// TwinCAT 3 PLC project TcoCognexVisionTests
// Title: TcoCognexVisionTests
// Company: Vortex.Library
// ProjectVersion: 0.6.0.913
// ProgramVersion: 3.1.4024.12
// libraries:
//   Tc2_Standard, * (Beckhoff Automation GmbH)
//   Tc2_System, * (Beckhoff Automation GmbH)
//   Tc3_Module, * (Beckhoff Automation GmbH)
//   TcoAbstractions, 0.6.0.913 (Vortex.Library)
//   TcoCognexVision, 0.6.0.913 (Vortex.Library)
//   TcoCore, 0.6.0.913 (Vortex.Library)
//   TcoInspectors, 0.6.0.913 (Vortex.Library)
//   TcoIo, 0.6.0.913 (Vortex.Library)
//   TcoUtilities, 0.6.0.913 (Vortex.Library)
// project tree:
//   DUTs/ DesignerResults.TcDUT, DesignerUserData.TcDUT
//   GVLs/ GVL.TcGVL
//   / PlcTask.TcTTO
//   POUs/ ITcoResultsData.TcIO, MAIN.TcPOU, myVeryFirstTcoContext.TcPOU, ProjectSpecificData.TcPOU
// (motion and I/O tree: see PLC project tcocognexvision)
// real-time tasks:
//   TASK PlcTask: cycle T#10ms, priority 20, ADS port 350
//   TASK PNIO: cycle T#16ms, priority 21, ADS port 351
//   TASK PlcTask1: cycle T#10ms, priority 22, ADS port 352
// variable links:
//   TcoCognexVisionTests/TcoCognexVisionTests Instance <-> Device 1 (Profinet Controller)/myveryfirstdataman
//     PlcTask Inputs/GVL.myVeryFirstDatamanGVL.AcquisitionStatus.Acquiring <-> API/Acquisition_Status/Acquisition_Status/Inputs/Acquisition_Status_Register/Acquiring
//     PlcTask Inputs/GVL.myVeryFirstDatamanGVL.AcquisitionStatus.MissedAcquisition <-> API/Acquisition_Status/Acquisition_Status/Inputs/Acquisition_Status_Register/Missed_Acquisition
//     PlcTask Inputs/GVL.myVeryFirstDatamanGVL.AcquisitionStatus.TriggerAcknowledge <-> API/Acquisition_Status/Acquisition_Status/Inputs/Acquisition_Status_Register/Trigger_Acknowledge
//     PlcTask Inputs/GVL.myVeryFirstDatamanGVL.AcquisitionStatus.TriggerID <-> API/Acquisition_Status/Acquisition_Status/Inputs/Trigger_ID
//     PlcTask Inputs/GVL.myVeryFirstDatamanGVL.AcquisitionStatus.TriggerReady <-> API/Acquisition_Status/Acquisition_Status/Inputs/Acquisition_Status_Register/Trigger_Ready
//     PlcTask Inputs/GVL.myVeryFirstDatamanGVL.PnIoBoxDiag <-> Inputs/PnIoBoxDiag
//     PlcTask Inputs/GVL.myVeryFirstDatamanGVL.PnIoBoxState <-> Inputs/PnIoBoxState
//     PlcTask Inputs/GVL.myVeryFirstDatamanGVL.ResultData.ResultCode <-> API/Result_Data_64_bytes/Result_Data_64_bytes/Inputs/Result_Code
//     PlcTask Inputs/GVL.myVeryFirstDatamanGVL.ResultData.ResultData <-> API/Result_Data_64_bytes/Result_Data_64_bytes/Inputs/Result_Data
//     PlcTask Inputs/GVL.myVeryFirstDatamanGVL.ResultData.ResultExtended <-> API/Result_Data_64_bytes/Result_Data_64_bytes/Inputs/Result_Extended
//     PlcTask Inputs/GVL.myVeryFirstDatamanGVL.ResultData.ResultID <-> API/Result_Data_64_bytes/Result_Data_64_bytes/Inputs/Result_ID
//     PlcTask Inputs/GVL.myVeryFirstDatamanGVL.ResultData.ResultLength <-> API/Result_Data_64_bytes/Result_Data_64_bytes/Inputs/Result_Length
//     PlcTask Inputs/GVL.myVeryFirstDatamanGVL.ResultsStatus.DecodeComplete <-> API/Results_Status/Results_Status/Inputs/Results_Status_Register/Decode_Complete
//     PlcTask Inputs/GVL.myVeryFirstDatamanGVL.ResultsStatus.Decoding <-> API/Results_Status/Results_Status/Inputs/Results_Status_Register/Decoding
//     PlcTask Inputs/GVL.myVeryFirstDatamanGVL.ResultsStatus.ErrorDetected <-> API/Results_Status/Results_Status/Inputs/Results_Status_Register/Set_when_reader_fault_occurs
//     PlcTask Inputs/GVL.myVeryFirstDatamanGVL.ResultsStatus.ResultsAvailable <-> API/Results_Status/Results_Status/Inputs/Results_Status_Register/Results_Available
//     PlcTask Inputs/GVL.myVeryFirstDatamanGVL.ResultsStatus.ResultsBufferOverrun <-> API/Results_Status/Results_Status/Inputs/Results_Status_Register/Results_Buffer_Overrun
//     PlcTask Inputs/GVL.myVeryFirstDatamanGVL.SoftEventControl.ExecuteDMCCAcknowledge <-> API/Soft_Event_Control/Soft_Event_Control/Inputs/Soft_Event_Acknowledge_Register/Execute_DMCC_Acknowledge
//     PlcTask Inputs/GVL.myVeryFirstDatamanGVL.SoftEventControl.SetMatchStringAcknowledge <-> API/Soft_Event_Control/Soft_Event_Control/Inputs/Soft_Event_Acknowledge_Register/Set_Match_String_Acknowledge
//     PlcTask Inputs/GVL.myVeryFirstDatamanGVL.SoftEventControl.TrainBrightnessAcknowledge <-> API/Soft_Event_Control/Soft_Event_Control/Inputs/Soft_Event_Acknowledge_Register/Train_Brightness_Acknowledge
//     PlcTask Inputs/GVL.myVeryFirstDatamanGVL.SoftEventControl.TrainCodeAcknowledge <-> API/Soft_Event_Control/Soft_Event_Control/Inputs/Soft_Event_Acknowledge_Register/Train_Code_Acknowledge
//     PlcTask Inputs/GVL.myVeryFirstDatamanGVL.SoftEventControl.TrainFocusAcknowledge <-> API/Soft_Event_Control/Soft_Event_Control/Inputs/Soft_Event_Acknowledge_Register/Train_Focus_Acknowledge
//     PlcTask Inputs/GVL.myVeryFirstDatamanGVL.SoftEventControl.TrainMatchStringAcknowledge <-> API/Soft_Event_Control/Soft_Event_Control/Inputs/Soft_Event_Acknowledge_Register/Train_Match_String_Acknowledge
//     PlcTask Inputs/GVL.myVeryFirstDatamanGVL.SoftEventControl.UntrainAcknowledge <-> API/Soft_Event_Control/Soft_Event_Control/Inputs/Soft_Event_Acknowledge_Register/Untrain_Acknowledge
//     PlcTask Outputs/GVL.myVeryFirstDatamanGVL.AcquisitionControl.Trigger <-> API/Acquisition_Control/Acquisition_Control/Outputs/Acquisition_Control_Register/Trigger
//     PlcTask Outputs/GVL.myVeryFirstDatamanGVL.AcquisitionControl.TriggerEnable <-> API/Acquisition_Control/Acquisition_Control/Outputs/Acquisition_Control_Register/Trigger_Enable
//     PlcTask Outputs/GVL.myVeryFirstDatamanGVL.PnIoBoxCtrl <-> Outputs/PnIoBoxCtrl
//     PlcTask Outputs/GVL.myVeryFirstDatamanGVL.ResultsControl.EnableResultBuffering <-> API/Results_Control/Results_Control/Outputs/Results_Control_Register/Enable_Result_Buffering
//     PlcTask Outputs/GVL.myVeryFirstDatamanGVL.ResultsControl.ResultsAcknowledge <-> API/Results_Control/Results_Control/Outputs/Results_Control_Register/Results_Acknowledge
//     PlcTask Outputs/GVL.myVeryFirstDatamanGVL.SoftEventControl.ExecuteDMCC <-> API/Soft_Event_Control/Soft_Event_Control/Outputs/Soft_Event_Control_Register/Execute_DMCC
//     PlcTask Outputs/GVL.myVeryFirstDatamanGVL.SoftEventControl.SetMatchString <-> API/Soft_Event_Control/Soft_Event_Control/Outputs/Soft_Event_Control_Register/Set_Match_String
//     PlcTask Outputs/GVL.myVeryFirstDatamanGVL.SoftEventControl.TrainBrightness <-> API/Soft_Event_Control/Soft_Event_Control/Outputs/Soft_Event_Control_Register/Train_Brightness
//     PlcTask Outputs/GVL.myVeryFirstDatamanGVL.SoftEventControl.TrainCode <-> API/Soft_Event_Control/Soft_Event_Control/Outputs/Soft_Event_Control_Register/Train_Code
//     PlcTask Outputs/GVL.myVeryFirstDatamanGVL.SoftEventControl.TrainFocus <-> API/Soft_Event_Control/Soft_Event_Control/Outputs/Soft_Event_Control_Register/Train_Focus
//     PlcTask Outputs/GVL.myVeryFirstDatamanGVL.SoftEventControl.TrainMatchString <-> API/Soft_Event_Control/Soft_Event_Control/Outputs/Soft_Event_Control_Register/Train_Match_String
//     PlcTask Outputs/GVL.myVeryFirstDatamanGVL.SoftEventControl.Untrain <-> API/Soft_Event_Control/Soft_Event_Control/Outputs/Soft_Event_Control_Register/Untrain
//     PlcTask Outputs/GVL.myVeryFirstDatamanGVL.UserData.UserData <-> API/User_Data_64_bytes/User_Data_64_bytes/Outputs/User_Data
//     PlcTask Outputs/GVL.myVeryFirstDatamanGVL.UserData.UserDataLength <-> API/User_Data_64_bytes/User_Data_64_bytes/Outputs/User_Data_Length
//     PlcTask Outputs/GVL.myVeryFirstDatamanGVL.UserData.UserDataOption <-> API/User_Data_64_bytes/User_Data_64_bytes/Outputs/User_Data_Option
//   TcoCognexVisionTests/TcoCognexVisionTests Instance <-> Device 1 (Profinet Controller)/myveryfirstinsight
//     PlcTask Inputs/GVL.myVeryFirstInsightGVL.AcquisitionStatus.AcquisitionID <-> API/Acquisition_Status/Acquisition_Status/Inputs/Acquisition_ID
//     PlcTask Inputs/GVL.myVeryFirstInsightGVL.AcquisitionStatus.AcquisitionTriggerAcknowledge <-> API/Acquisition_Status/Acquisition_Status/Inputs/Acquisition_Status_Register/Acquisition_Trigger_Acknowledge
//     PlcTask Inputs/GVL.myVeryFirstInsightGVL.AcquisitionStatus.AcquisitionTriggerReady <-> API/Acquisition_Status/Acquisition_Status/Inputs/Acquisition_Status_Register/Acquisition_Trigger_Ready
//     PlcTask Inputs/GVL.myVeryFirstInsightGVL.AcquisitionStatus.ExposureComplete <-> API/Acquisition_Status/Acquisition_Status/Inputs/Acquisition_Status_Register/Exposure_Complete
//     PlcTask Inputs/GVL.myVeryFirstInsightGVL.AcquisitionStatus.MissedAcquisition <-> API/Acquisition_Status/Acquisition_Status/Inputs/Acquisition_Status_Register/Missed_Acquisition
//     PlcTask Inputs/GVL.myVeryFirstInsightGVL.AcquisitionStatus.OfflineReason0 <-> API/Acquisition_Status/Acquisition_Status/Inputs/Acquisition_Status_Register/Offline_Reason_0
//     PlcTask Inputs/GVL.myVeryFirstInsightGVL.AcquisitionStatus.OfflineReason1 <-> API/Acquisition_Status/Acquisition_Status/Inputs/Acquisition_Status_Register/Offline_Reason_1
//     PlcTask Inputs/GVL.myVeryFirstInsightGVL.AcquisitionStatus.OfflineReason2 <-> API/Acquisition_Status/Acquisition_Status/Inputs/Acquisition_Status_Register/Offline_Reason_2
//     PlcTask Inputs/GVL.myVeryFirstInsightGVL.AcquisitionStatus.Online <-> API/Acquisition_Status/Acquisition_Status/Inputs/Acquisition_Status_Register/Online
//     PlcTask Inputs/GVL.myVeryFirstInsightGVL.CommandControl.CurrentJobID <-> API/Command_Control/Command_Control/Inputs/Current_Job_ID
//     PlcTask Inputs/GVL.myVeryFirstInsightGVL.InspectionStatus.CommandComplete <-> API/Inspection_Status/Inspection_Status/Inputs/Inspection_Status_Register/Command_Complete
//     PlcTask Inputs/GVL.myVeryFirstInsightGVL.InspectionStatus.CommandExecuting <-> API/Inspection_Status/Inspection_Status/Inputs/Inspection_Status_Register/Command_Executing
//     PlcTask Inputs/GVL.myVeryFirstInsightGVL.InspectionStatus.CommandFailed <-> API/Inspection_Status/Inspection_Status/Inputs/Inspection_Status_Register/Command_Failed
//     PlcTask Inputs/GVL.myVeryFirstInsightGVL.InspectionStatus.Error <-> API/Inspection_Status/Inspection_Status/Inputs/Inspection_Status_Register/Error
//     PlcTask Inputs/GVL.myVeryFirstInsightGVL.InspectionStatus.ErrorCode <-> API/Inspection_Status/Inspection_Status/Inputs/Error_Code
//     PlcTask Inputs/GVL.myVeryFirstInsightGVL.InspectionStatus.ExtendedUserDataSetAcknowledge <-> API/Inspection_Status/Inspection_Status/Inputs/Inspection_Status_Register/Extended_User_Data_Set_Acknowledge
//     PlcTask Inputs/GVL.myVeryFirstInsightGVL.InspectionStatus.InspectionCompleted <-> API/Inspection_Status/Inspection_Status/Inputs/Inspection_Status_Register/Inspection_Completed
//     PlcTask Inputs/GVL.myVeryFirstInsightGVL.InspectionStatus.OverallJobPassFail <-> API/Inspection_Status/Inspection_Status/Inputs/Inspection_Status_Register/Set_when_last_inspection_passed,_based_on_the_Overall_Job_Pass_Fail_cell
//     PlcTask Inputs/GVL.myVeryFirstInsightGVL.InspectionStatus.ResultsBufferOverrun <-> API/Inspection_Status/Inspection_Status/Inputs/Inspection_Status_Register/Results_Buffer_Overrun
//     PlcTask Inputs/GVL.myVeryFirstInsightGVL.InspectionStatus.ResultsValid <-> API/Inspection_Status/Inspection_Status/Inputs/Inspection_Status_Register/Results_Valid
//     PlcTask Inputs/GVL.myVeryFirstInsightGVL.InspectionStatus.SystemBusy <-> API/Inspection_Status/Inspection_Status/Inputs/Inspection_Status_Register/System_Busy
//     PlcTask Inputs/GVL.myVeryFirstInsightGVL.InspectionStatus.TestRunReady <-> API/Inspection_Status/Inspection_Status/Inputs/Inspection_Status_Register/Test_Run_Ready
//     PlcTask Inputs/GVL.myVeryFirstInsightGVL.PnIoBoxDiag <-> Inputs/PnIoBoxDiag
//     PlcTask Inputs/GVL.myVeryFirstInsightGVL.PnIoBoxState <-> Inputs/PnIoBoxState
//     PlcTask Inputs/GVL.myVeryFirstInsightGVL.ResultsData.InspectionID <-> API/Results_128_bytes/Results_128_bytes/Inputs/Inspection ID
//     PlcTask Inputs/GVL.myVeryFirstInsightGVL.ResultsData.InspectionResults <-> API/Results_128_bytes/Results_128_bytes/Inputs/Inspection Results
//     PlcTask Inputs/GVL.myVeryFirstInsightGVL.ResultsData.ResultCode <-> API/Results_128_bytes/Results_128_bytes/Inputs/Result Code
//     PlcTask Inputs/GVL.myVeryFirstInsightGVL.SoftEventControl.TriggerSoftEventAcknowledge[{0..7}] <-> API/SoftEvent_Control/SoftEvent_Control/Inputs/SoftEvent_Status/Trigger_SoftEvent_{0..7}_Acknowledge  (8 links)
//     PlcTask Outputs/GVL.myVeryFirstInsightGVL.AcquisitionControl.AcquisitionTrigger <-> API/Acquisition_Control/Acquisition_Control/Outputs/Acquisition_Control_Register/Acquisition_Trigger
//     PlcTask Outputs/GVL.myVeryFirstInsightGVL.AcquisitionControl.AcquisitionTriggerEnable <-> API/Acquisition_Control/Acquisition_Control/Outputs/Acquisition_Control_Register/Acquisition_Trigger_Enable
//     PlcTask Outputs/GVL.myVeryFirstInsightGVL.AcquisitionControl.ClearExposureComplete <-> API/Acquisition_Control/Acquisition_Control/Outputs/Acquisition_Control_Register/Clear_Exposure_Complete
//     PlcTask Outputs/GVL.myVeryFirstInsightGVL.AcquisitionControl.SetOffline <-> API/Acquisition_Control/Acquisition_Control/Outputs/Acquisition_Control_Register/Set_Offline
//     PlcTask Outputs/GVL.myVeryFirstInsightGVL.CommandControl.Command <-> API/Command_Control/Command_Control/Outputs/Command
//     PlcTask Outputs/GVL.myVeryFirstInsightGVL.InspectionControl.AcknowledgeInspectionResults <-> API/Inspection_Control/Inspection_Control/Outputs/Inspection_Control_Register/Acknowledge_Inspection_Results
//     PlcTask Outputs/GVL.myVeryFirstInsightGVL.InspectionControl.ClearError <-> API/Inspection_Control/Inspection_Control/Outputs/Inspection_Control_Register/Clear_Error
//     PlcTask Outputs/GVL.myVeryFirstInsightGVL.InspectionControl.EnableResultsBuffering <-> API/Inspection_Control/Inspection_Control/Outputs/Inspection_Control_Register/Enable_Results_Buffering
//     PlcTask Outputs/GVL.myVeryFirstInsightGVL.InspectionControl.ExecuteCommand <-> API/Inspection_Control/Inspection_Control/Outputs/Inspection_Control_Register/Execute_Command
//     PlcTask Outputs/GVL.myVeryFirstInsightGVL.InspectionControl.ExtendedUserDataSet <-> API/Inspection_Control/Inspection_Control/Outputs/Inspection_Control_Register/Extended_User_Data_Set
//     PlcTask Outputs/GVL.myVeryFirstInsightGVL.PnIoBoxCtrl <-> Outputs/PnIoBoxCtrl
//     PlcTask Outputs/GVL.myVeryFirstInsightGVL.SoftEventControl.TriggerSoftEvent[{0..7}] <-> API/SoftEvent_Control/SoftEvent_Control/Outputs/SoftEvent_Control/Trigger_SoftEvent_{0..7}  (8 links)
//     PlcTask Outputs/GVL.myVeryFirstInsightGVL.UserData.UserData <-> API/User_Data_128_bytes/User_Data_128 bytes/Outputs/User Data

CONFIGURATION TcoCognexVisionTests
    RESOURCE PLC ON TwinCAT3
        TASK PlcTask(INTERVAL := T#16ms, PRIORITY := 21);
        PROGRAM MAIN WITH PlcTask : MAIN;
    END_RESOURCE
END_CONFIGURATION

// ---- DUTs/DesignerResults.TcDUT
TYPE DesignerResults EXTENDS TcoCore.TcoStruct :
STRUCT
	{attribute addProperty Name "<#ResultBool#>"}
	ResultBool:BOOL;
	{attribute addProperty Name "<#ResultInt#>"}
	ResultInt:INT;
	{attribute addProperty Name "<#ResultString#>"}
	ResultString:STRING;

	
	{attribute addProperty Name "<#Data inspector#>"}
	DigitalInspector:TcoInspectors.TcoDigitalInspector(THISSTRUCT);
	{attribute addProperty Name "<#Data inspector#>"}
	DataInspector:TcoInspectors.TcoDataInspector(THISSTRUCT);
	
	{attribute addProperty Name "<#Analog inspector#>"}
	AnalogInspector:TcoInspectors.TcoAnalogueInspector(THISSTRUCT);
END_STRUCT
END_TYPE

// ---- DUTs/DesignerUserData.TcDUT
TYPE DesignerUserData EXTENDS TcoCore.TcoStruct :
STRUCT
	{attribute addProperty Name "<#ResultBool#>"}
	ResultBool:BOOL;
	{attribute addProperty Name "<#ResultInt#>"}
	ResultInt:INT;
	{attribute addProperty Name "<#ResultString#>"}
	ResultString:STRING;
	
END_STRUCT
END_TYPE

// ---- GVLs/GVL.TcGVL
{attribute 'qualified_only'}
VAR_GLOBAL
	myVeryFirstDatamanGVL 	: TcoCognexVision.TcoDatamanIO_v_5_x_x;
	myVeryFirstInsightGVL 	: TcoCognexVision.TcoInsightIO_v_5_x_x;
END_VAR

// ---- POUs/ITcoResultsData.TcIO
INTERFACE ITcoResultsData

END_INTERFACE

// ---- POUs/MAIN.TcPOU
PROGRAM MAIN
VAR
	myVeryFirstTcoContextInstance :	myVeryFirstTcoContext;
END_VAR

myVeryFirstTcoContextInstance.Run();

END_PROGRAM

// ---- POUs/myVeryFirstTcoContext.TcPOU
FUNCTION_BLOCK myVeryFirstTcoContext EXTENDS TcoCore.TcoContext
VAR
	{attribute addProperty Name "<#My very first DATAMAN#>"}
	myVeryFirstDataman : TcoCognexVision.TcoDataman_v_5_x_x(THIS^);
	{attribute addProperty Name "<#My very first INSIGHT#>"}
	myVeryFirstInsight : TcoCognexVision.TcoInsight_v_5_x_x(THIS^);

	

	{attribute addProperty Name "<#Cognex Designer#>"}
	designer : TcoCognexVision.TcoDesigner_v_2_x_x(THIS^);
	
	{attribute addProperty Name "<#Project Specific Data#>"}
    _specificData : ProjectSpecificData(THIS^);
	
	

END_VAR

(*~
	<docu>
		<summary>
			Main method of the TcoContext. This is the entry point of any control logic that belongs to this context. 
			The call of this method is ensured by calling the <c>InstanceName.Run()</c> method, and it must not be called explicitly.
			This method is abstract, and it must be overridden in derived block.
		</summary>
	</docu>
~*)
METHOD PROTECTED  Main

VAR
	
END_VAR
myVeryFirstDataman(inoIoData:= GVL.myVeryFirstDatamanGVL);
myVeryFirstDataman.Service();

myVeryFirstInsight.Config.UserDataSize := eTcoInsightUserDataSize_v_5_x_x.USER_DATA_128B;
myVeryFirstInsight.Config.ResultDataSize := eTcoInsightResultDataSize_v_5_x_x.RESULT_DATA_128B;
myVeryFirstInsight(inoIoData:= GVL.myVeryFirstInsightGVL);
myVeryFirstInsight.Service();
myVeryFirstDataman.Read();
myVeryFirstDataman.GetResultAsString(0,myVeryFirstDataman.Status.SignalStatus.ResultLength);




designer(inoData:=_specificData );
designer.Service();
END_METHOD

END_FUNCTION_BLOCK

// ---- POUs/ProjectSpecificData.TcPOU
FUNCTION_BLOCK ProjectSpecificData EXTENDS TcoCognexVision.TcoDesignerRootContainer  
VAR_INPUT
END_VAR
VAR_OUTPUT
END_VAR
VAR
	{attribute wpf [Container(Layout.Stack,"PcToPlc")]}	
	{attribute wpf [Group(Layout.GroupBox)]}
	{attribute addProperty Name "<#PcToPlc#>"}
	PcToPlc:DesignerResults;
	{attribute wpf [Container(Layout.Stack,"PlcToPc")]}	
	{attribute wpf [Group(Layout.GroupBox)]}
	{attribute addProperty Name "<#PlcToPc#>"}
	PlcToPc:DesignerUserData;
	
END_VAR

PROPERTY PUBLIC Results : REFERENCE TO DesignerResults
GET
Results ref= PcToPlc;
END_GET
END_PROPERTY

PROPERTY PUBLIC UserData : REFERENCE TO DesignerUserData
GET
UserData ref= PlcToPc;
END_GET
END_PROPERTY

END_FUNCTION_BLOCK
